// TIA Portal V21 export
FUNCTION "FC_FillHelper" : Real   // FC7, SCL
TITLE = Volume from raw flow
// Unpublished helper of the filling unit
// stored: Namespace Filling, SetENOAutomatically false
   VAR_INPUT
      RawFlow : Int;   // Raw flow value
      Factor : Real;   // Litres per raw unit
   END_VAR
BEGIN

       #FC_FillHelper := INT_TO_REAL(#RawFlow) * #Factor;
END_FUNCTION
